// Axis the operator jogs in manual mode.
{attribute 'qualified_only'}
{attribute 'strict'}
TYPE E_JogAxis :
(
    eTravel := 0,
    eHoist  := 1,
    eFork   := 2
) INT;
END_TYPE

(* stored: Version 1.1.0.1
   DUT E_JogAxis: Id {84e3cc36-13e1-045d-34c6-93772e773ecc} *)
